Fanuc KAREL source: kt00039.KL

-- PROVISIONAL review KL for V1013-1; original PC SHA256 055e80f32aa04b58b7e91d7c96a0978f4faae2e700b49855c7e97bd0665c9b2d
-- Incomplete behavior may be omitted. Consult companion uncertainty JSON. Do not deploy.
PROGRAM KT00039
%NOLOCKGROUP
VAR
  I1 : INTEGER
  OUT : INTEGER
-- UNRESOLVED_DECL H2 type=002017
BEGIN
  -- UNRESOLVED_PC offsets 5-16; opcodes 2E,23
  -- UNRESOLVED_PC offsets 21-35; opcodes 2E,22,9D,33,B4
  -- UNRESOLVED_PC offsets 40-62; opcodes 21,22,9D,33,B3,53,23
  -- UNRESOLVED_PC offsets 67-71; opcodes 7F
END KT00039
